(* IEC 61131-3 sources: avi-aoi-management/server/services/programming/iec61131/golden-st/valid, 35 files *)

(* ---- v01-probe-fb.st ---- *)
FUNCTION_BLOCK FB_Light
VAR_INPUT
  Enable : BOOL;
END_VAR
VAR_OUTPUT
  Red : BOOL;
END_VAR
VAR
  T1 : TON;
END_VAR
Red := Enable;
END_FUNCTION_BLOCK

(* ---- v11-fb-in-out-temp-instance.st ---- *)
FUNCTION_BLOCK FB_Accumulate
VAR_INPUT
    Add    : REAL;
    Enable : BOOL;
END_VAR
VAR_IN_OUT
    Total : REAL;
END_VAR
VAR_OUTPUT
    Overflow : BOOL;
END_VAR
VAR_TEMP
    Tmp : REAL;
END_VAR
VAR CONSTANT
    LIMIT_MAX : REAL := 1.0E6;
END_VAR
    IF Enable THEN
        Tmp := Total + Add;
        Overflow := Tmp > LIMIT_MAX;
        IF NOT Overflow THEN
            Total := Tmp;
        END_IF;
    END_IF;
END_FUNCTION_BLOCK

PROGRAM Main
VAR
    Acc     : FB_Accumulate;
    Energy  : REAL;
    Alarm   : BOOL;
END_VAR
    Acc(Add := 0.5, Enable := TRUE, Total := Energy);
    Alarm := Acc.Overflow;
END_PROGRAM

(* ---- v23-traffic-light-fb-timer-array.st ---- *)
FUNCTION_BLOCK FB_TrafficLight
VAR_INPUT
    Enable : BOOL;
END_VAR
VAR_OUTPUT
    Red    : BOOL;
    Yellow : BOOL;
    Green  : BOOL;
END_VAR
VAR
    Phase  : INT := 0;
    Timers : ARRAY[0..2] OF TON;
    Times  : ARRAY[0..2] OF TIME := [T#10s, T#3s, T#8s];
END_VAR

IF NOT Enable THEN
    Phase := 0;
    Red := TRUE; Yellow := FALSE; Green := FALSE;
    RETURN;
END_IF;

Timers[Phase](IN := TRUE, PT := Times[Phase]);
IF Timers[Phase].Q THEN
    Timers[Phase](IN := FALSE);
    Phase := (Phase + 1) MOD 3;
END_IF;

Red := Phase = 0;
Green := Phase = 1;
Yellow := Phase = 2;

END_FUNCTION_BLOCK

PROGRAM Crossing
VAR
    Light : FB_TrafficLight;
    Run   : BOOL := TRUE;
    Stop  : BOOL;
END_VAR
Light(Enable := Run);
Stop := Light.Red;
END_PROGRAM

(* ---- v25-std-functions-conversions.st ---- *)
FUNCTION_BLOCK FB_Clamp
VAR_INPUT
    In   : REAL;
    Lo   : REAL := 0.0;
    Hi   : REAL := 100.0;
END_VAR
VAR_OUTPUT
    Out     : REAL;
    Clipped : BOOL;
    Rounded : INT;
END_VAR
    Out := LIMIT(Lo, In, Hi);
    Clipped := Out <> In;
    Rounded := REAL_TO_INT(Out);
    Rounded := TRUNC(Out);
    Out := MAX(Out, INT_TO_REAL(Rounded));
END_FUNCTION_BLOCK

PROGRAM UseClamp
VAR
    Clamp : FB_Clamp;
    Raw   : REAL;
    Value : REAL;
    Warn  : BOOL;
END_VAR
    Clamp(In := Raw, Hi := 80.0, Out => Value, Clipped => Warn);
END_PROGRAM

(* ---- v32-r-edge-f-edge-inputs.st ---- *)
FUNCTION_BLOCK FB_EdgeCounter
VAR_INPUT
    Pulse   : BOOL R_EDGE;
    Release : BOOL F_EDGE;
    Reset   : BOOL;
END_VAR
VAR_OUTPUT
    Rising  : INT;
    Falling : INT;
END_VAR
IF Reset THEN
    Rising := 0;
    Falling := 0;
END_IF;
IF Pulse THEN
    Rising := Rising + 1;
END_IF;
IF Release THEN
    Falling := Falling + 1;
END_IF;
END_FUNCTION_BLOCK

PROGRAM UseEdges
VAR
    Counter : FB_EdgeCounter;
    Sensor  : BOOL;
    Total   : INT;
END_VAR
Counter(Pulse := Sensor, Release := Sensor, Reset := FALSE);
Total := Counter.Rising;
END_PROGRAM

(* ---- v02-probe-cmt.st ---- *)
PROGRAM P
VAR
  a : BOOL;
END_VAR
(* turn on if sensor is on *)
a := TRUE;
END_PROGRAM

(* ---- v03-conveyor-start-stop-ton.st ---- *)
(* Conveyor: Start push-button latches the motor, NC Stop drops it,
   a TON delays the running lamp by 2 s. *)
PROGRAM ConveyorStartStop
VAR_INPUT
    StartPB   : BOOL;          (* NO push-button *)
    StopPB_NC : BOOL := TRUE;  (* NC push-button: FALSE when pressed *)
END_VAR
VAR_OUTPUT
    Motor      : BOOL;
    RunningLmp : BOOL;
END_VAR
VAR
    RunDelay : TON;
END_VAR

Motor := (StartPB OR Motor) AND StopPB_NC;
RunDelay(IN := Motor, PT := T#2s);
RunningLmp := RunDelay.Q;

END_PROGRAM

(* ---- v04-debounce-ton.st ---- *)
PROGRAM DebounceInputSignal
VAR
    RawSignal    : BOOL;             (* noisy field input *)
    DebounceTmr  : TON;              (* standard on-delay timer instance *)
    StableSignal : BOOL;             (* debounced, steady result (output) *)
    DebounceTime : TIME := T#20ms;   (* dwell needed to accept a change *)
END_VAR

(* TON keeps Q low until IN has stayed high past PT (DebounceTime);
   this rejects contact chatter on a mechanical input. *)
DebounceTmr(IN := RawSignal, PT := DebounceTime);
StableSignal := DebounceTmr.Q;

END_PROGRAM

(* ---- v05-moving-average-array-for.st ---- *)
PROGRAM MovingAverage
VAR
    Samples    : ARRAY[0..7] OF REAL;
    WriteIndex : INT := 0;
    Idx        : INT;
    Sum        : REAL := 0.0;
    NewSample  : REAL;
    Average    : REAL;
END_VAR

Samples[WriteIndex] := NewSample;
WriteIndex := WriteIndex + 1;
IF WriteIndex >= 8 THEN
    WriteIndex := 0;
END_IF;

Sum := 0.0;
FOR Idx := 0 TO 7 DO
    Sum := Sum + Samples[Idx];
END_FOR;
Average := Sum / 8.0;

END_PROGRAM

(* ---- v06-case-enum-state-machine.st ---- *)
TYPE
    E_FillState : (Idle, Filling, Settling, Done);
END_TYPE

PROGRAM FillStation
VAR
    State      : E_FillState := Idle;
    StartReq   : BOOL;
    LevelHigh  : BOOL;
    Valve      : BOOL;
    SettleTmr  : TON;
END_VAR

CASE State OF
    Idle:
        Valve := FALSE;
        IF StartReq THEN
            State := Filling;
        END_IF;
    Filling:
        Valve := TRUE;
        IF LevelHigh THEN
            State := E_FillState#Settling;
        END_IF;
    Settling:
        Valve := FALSE;
        SettleTmr(IN := TRUE, PT := T#3s);
        IF SettleTmr.Q THEN
            SettleTmr(IN := FALSE);
            State := Done;
        END_IF;
    Done:
        IF NOT StartReq THEN
            State := Idle;
        END_IF;
END_CASE;

END_PROGRAM

(* ---- v07-case-int-ranges-else.st ---- *)
PROGRAM SpeedSelector
VAR
    Mode     : INT;
    SpeedSet : REAL;
    Fault    : BOOL;
END_VAR

CASE Mode OF
    0:
        SpeedSet := 0.0;
    1, 2:
        SpeedSet := 25.0;
    3..5:
        SpeedSet := 50.0 + INT_TO_REAL(Mode) * 5.0;
ELSE
    SpeedSet := 0.0;
    Fault := TRUE;
END_CASE

END_PROGRAM

(* ---- v08-while-exit.st ---- *)
PROGRAM FindFirstEmpty
VAR
    Slots     : ARRAY[1..10] OF BOOL;
    I         : INT;
    FirstFree : INT := -1;
END_VAR

I := 1;
WHILE I <= 10 DO
    IF NOT Slots[I] THEN
        FirstFree := I;
        EXIT;
    END_IF;
    I := I + 1;
END_WHILE;

END_PROGRAM

(* ---- v09-repeat-until.st ---- *)
PROGRAM ShiftRegister
VAR
    Reg   : ARRAY[0..4] OF INT;
    K     : INT;
    Input : INT;
END_VAR

K := 4;
REPEAT
    Reg[K] := Reg[K - 1];
    K := K - 1;
UNTIL K = 0
END_REPEAT;
Reg[0] := Input;

END_PROGRAM

(* ---- v10-function-var-input.st ---- *)
FUNCTION Scale : REAL
VAR_INPUT
    Raw    : INT;
    RawMax : INT;
    EngMax : REAL;
END_VAR
    IF RawMax <= 0 THEN
        Scale := 0.0;
        RETURN;
    END_IF;
    Scale := INT_TO_REAL(Raw) / INT_TO_REAL(RawMax) * EngMax;
END_FUNCTION

PROGRAM Main
VAR
    AnalogIn : INT;
    Pressure : REAL;
END_VAR
    Pressure := Scale(Raw := AnalogIn, RawMax := 27648, EngMax := 10.0);
    Pressure := Scale(AnalogIn, 27648, 16.0);
END_PROGRAM

(* ---- v12-ctu-rtrig-batch.st ---- *)
PROGRAM BatchCounter
VAR
    PartSensor : BOOL;
    ResetPB    : BOOL;
    Edge       : R_TRIG;
    Counter    : CTU;
    BatchDone  : BOOL;
    Count      : INT;
END_VAR

Edge(CLK := PartSensor);
Counter(CU := Edge.Q, R := ResetPB, PV := 50);
BatchDone := Counter.Q;
Count := Counter.CV;

END_PROGRAM

(* ---- v13-ctud-ctd.st ---- *)
PROGRAM BufferLevel
VAR
    InSensor  : BOOL;
    OutSensor : BOOL;
    Clear     : BOOL;
    Load      : BOOL;
    Level     : CTUD;
    Remaining : CTD;
    Full      : BOOL;
    Empty     : BOOL;
    Parts     : INT;
END_VAR

Level(CU := InSensor, CD := OutSensor, R := Clear, LD := FALSE, PV := 20);
Full := Level.QU;
Empty := Level.QD;
Parts := Level.CV;
Remaining(CD := OutSensor, LD := Load, PV := 100);
IF Remaining.Q THEN
    Load := TRUE;
END_IF;

END_PROGRAM

(* ---- v14-sr-rs-ftrig.st ---- *)
PROGRAM Latches
VAR
    SetBtn    : BOOL;
    ResetBtn  : BOOL;
    Released  : F_TRIG;
    PumpLatch : SR;
    FanLatch  : RS;
    Pump      : BOOL;
    Fan       : BOOL;
END_VAR

Released(CLK := SetBtn);
PumpLatch(S1 := SetBtn, R := ResetBtn);
FanLatch(S := Released.Q, R1 := ResetBtn);
Pump := PumpLatch.Q1;
Fan := FanLatch.Q1;

END_PROGRAM

(* ---- v15-struct-members.st ---- *)
TYPE
    ST_Axis : STRUCT
        Position : REAL;
        Velocity : REAL;
        Homed    : BOOL;
    END_STRUCT;
    ST_Cell : STRUCT
        AxisX : ST_Axis;
        AxisY : ST_Axis;
        Name  : STRING[32];
    END_STRUCT;
END_TYPE

PROGRAM CellStatus
VAR
    Cell     : ST_Cell;
    AllHomed : BOOL;
    Dist     : REAL;
END_VAR

AllHomed := Cell.AxisX.Homed AND Cell.AxisY.Homed;
Dist := SQRT(Cell.AxisX.Position * Cell.AxisX.Position + Cell.AxisY.Position ** 2.0);
Cell.Name := 'Cell A';

END_PROGRAM

(* ---- v16-comments-with-keywords.st ---- *)
// if this line were code it would be broken: IF x THEN
(* Multi-line comment mentioning for, while, repeat and END_IF / END_FOR
   and even an unbalanced VAR or two: VAR VAR VAR *)
PROGRAM CommentTorture
VAR
    Lamp  : BOOL;   // turn on if the door is open
    Door  : BOOL;   (* while door open, for safety keep lamp on *)
    Label : STRING := 'IF Door THEN END_WHILE (* not a comment *)';
END_VAR
/* block comment: FOR i := 1 TO 10 DO */
IF Door THEN   // for the operator
    Lamp := TRUE;  (* end_if would go here if *)
ELSE
    Lamp := FALSE;
END_IF;
Label := 'it$'s $'quoted$' and // not a comment';
END_PROGRAM

(* ---- v17-global-external-retain.st ---- *)
VAR_GLOBAL
    gMachineReady : BOOL;
    gCycleCount   : DINT;
END_VAR

PROGRAM Cycle
VAR_EXTERNAL
    gMachineReady : BOOL;
    gCycleCount   : DINT;
END_VAR
VAR RETAIN
    TotalCycles : DINT;
END_VAR
VAR CONSTANT
    MAX_CYCLES : DINT := 1000000;
END_VAR
VAR
    CycleStart : BOOL;
    Edge       : R_TRIG;
END_VAR

Edge(CLK := CycleStart AND gMachineReady);
IF Edge.Q AND (TotalCycles < MAX_CYCLES) THEN
    TotalCycles := TotalCycles + 1;
    gCycleCount := TotalCycles;
END_IF;

END_PROGRAM

(* ---- v18-typed-literals.st ---- *)
PROGRAM Literals
VAR
    Mask     : WORD := 16#00FF;
    Bits     : BYTE := 2#1010_0101;
    Oct      : INT := 8#17;
    Small    : INT := INT#5;
    Big      : DINT := 1_000_000;
    Sci      : LREAL := 1.5E-3;
    Neg      : INT := -42;
    Dwell    : TIME := T#1h2m3s;
    Short    : TIME := TIME#500ms;
    Frac     : TIME := T#1.5s;
    Day      : DATE := D#2024-01-31;
    Clock    : TOD := TOD#12:30:00;
    Stamp    : DT := DT#2024-01-31-08:15:00;
    Flag     : BOOL := BOOL#TRUE;
    Masked   : WORD;
END_VAR

Masked := Mask AND 16#0F0F;
IF Dwell > T#1h THEN
    Flag := FALSE;
END_IF;

END_PROGRAM

(* ---- v19-direct-addresses.st ---- *)
PROGRAM IoMapping
VAR
    StartBtn AT %IX0.0 : BOOL;
    StopBtn  AT %IX0.1 : BOOL;
    Motor    AT %QX0.0 : BOOL;
    Speed    AT %IW0   : INT;
    SpeedOut AT %QW0   : INT;
END_VAR

Motor := StartBtn AND NOT StopBtn;
SpeedOut := Speed;
%QX0.1 := Motor;
%MW10 := Speed / 2;

END_PROGRAM

(* ---- v20-expressions-operators.st ---- *)
PROGRAM Expressions
VAR
    A, B, C : BOOL;
    X, Y    : INT;
    R       : REAL;
    Res     : BOOL;
    Parity  : INT;
END_VAR

Res := (A AND B) OR (NOT C XOR A) & (X <> Y);
Res := (X >= 10) AND (Y <= -3) OR (X = Y) AND NOT (X > Y OR X < Y);
Parity := X MOD 2;
R := INT_TO_REAL(X) ** 2.0 + INT_TO_REAL(Y) / 3.0 - 1.0;
X := -(Y * 4) + ABS(Y) - MAX(X, Y) + MIN(X, 0) + LIMIT(0, Y, 100);
Res := SEL(A, B, C);

END_PROGRAM

(* ---- v21-fb-output-binding.st ---- *)
PROGRAM OutputBinding
VAR
    Go       : BOOL;
    Tmr      : TON;
    Done     : BOOL;
    Elapsed  : TIME;
    Pulse    : TP;
    OffDelay : TOF;
    PulseOut : BOOL;
    Hold     : BOOL;
END_VAR

Tmr(IN := Go, PT := T#2s, Q => Done, ET => Elapsed);
Pulse(IN := Done, PT := T#500ms, Q => PulseOut);
OffDelay(IN := Go, PT := T#5s);
Hold := OffDelay.Q AND NOT Pulse.Q;

END_PROGRAM

(* ---- v22-nested-if-for-by.st ---- *)
PROGRAM Nested
VAR
    Data  : ARRAY[1..20] OF INT;
    I     : INT;
    Pos   : INT;
    Neg   : INT;
    Zero  : INT;
END_VAR

Pos := 0; Neg := 0; Zero := 0;
FOR I := 20 TO 1 BY -1 DO
    IF Data[I] > 0 THEN
        Pos := Pos + 1;
    ELSIF Data[I] < 0 THEN
        Neg := Neg + 1;
        IF Neg > 5 THEN
            EXIT;
        END_IF;
    ELSE
        Zero := Zero + 1;
    END_IF;
END_FOR;

END_PROGRAM

(* ---- v24-strings-bits-multidim.st ---- *)
PROGRAM StringsAndBits
VAR
    Status  : WORD;
    Ready   : BOOL;
    Msg     : STRING(80);
    Prefix  : STRING := 'Line';
    Grid    : ARRAY[1..3, 1..4] OF INT;
    MsgLen  : INT;
    R, C    : INT;
END_VAR

Ready := Status.3;
Status.0 := TRUE;
Msg := CONCAT(Prefix, ' 1 ready');
MsgLen := LEN(Msg);
FOR R := 1 TO 3 DO
    FOR C := 1 TO 4 DO
        Grid[R, C] := R * 10 + C;
    END_FOR;
END_FOR;

END_PROGRAM

(* ---- v26-unbounded-while-lint-only.st ---- *)
(* Syntactically valid; the SAFETY linter (not the parser) flags the unbounded loop. *)
PROGRAM ConveyorPoll
VAR
    SensorInput : BOOL;
    MotorRun    : BOOL;
END_VAR

WHILE TRUE DO
    MotorRun := SensorInput;
END_WHILE;

END_PROGRAM

(* ---- v27-time-date-functions.st ---- *)
PROGRAM TimeArithmetic
VAR
    Dwell     : TIME := T#2s;
    Extra     : TIME := T#500ms;
    Total     : TIME;
    Diff      : TIME;
    Scaled    : TIME;
    Half      : TIME;
    ShiftTod  : TOD := TOD#06:00:00;
    NowTod    : TOD := TOD#14:30:00;
    LaterTod  : TOD;
    EarlyTod  : TOD;
    Stamp     : DT := DT#2024-01-31-08:15:00;
    Stamp2    : DT;
    Stamp3    : DT;
    Day1      : DATE := D#2024-01-01;
    Day2      : DATE := D#2024-02-01;
    DaySpan   : TIME;
    TodSpan   : TIME;
    DtSpan    : TIME;
    Joined    : DT;
END_VAR

Total := ADD_TIME(Dwell, Extra);
Diff := SUB_TIME(Dwell, Extra);
Scaled := MULTIME(Dwell, 3);
Half := DIVTIME(Dwell, 2);
LaterTod := ADD_TOD_TIME(ShiftTod, T#8h);
EarlyTod := SUB_TOD_TIME(NowTod, T#30m);
TodSpan := SUB_TOD_TOD(NowTod, ShiftTod);
Stamp2 := ADD_DT_TIME(Stamp, T#1h);
Stamp3 := SUB_DT_TIME(Stamp, T#15m);
DtSpan := SUB_DT_DT(Stamp2, Stamp);
DaySpan := SUB_DATE_DATE(Day2, Day1);
Joined := CONCAT_DATE_TOD(Day1, ShiftTod);

END_PROGRAM

(* ---- v28-long-conversions-bcd.st ---- *)
PROGRAM Conversions
VAR
    Stamp    : DATE_AND_TIME := DT#2024-01-31-08:15:00;
    ClockTod : TIME_OF_DAY;
    OnlyDay  : DATE;
    Raw      : WORD := 16#0123;
    Value    : INT;
    Back     : WORD;
    R        : REAL := 12.7;
    I        : DINT;
    Text     : STRING;
    B        : BOOL;
END_VAR

ClockTod := DATE_AND_TIME_TO_TIME_OF_DAY(Stamp);
OnlyDay := DATE_AND_TIME_TO_DATE(Stamp);
ClockTod := DT_TO_TOD(Stamp);
Value := WORD_BCD_TO_INT(Raw);
Value := BCD_TO_INT(Raw);
Back := INT_TO_BCD(Value);
I := REAL_TO_DINT(R);
I := TRUNC(R);
Text := INT_TO_STRING(Value);
B := INT_TO_BOOL(Value);

END_PROGRAM

(* ---- v29-numeric-selection-shift.st ---- *)
PROGRAM NumericSelectShift
VAR
    X, Y, Z  : REAL;
    A, B     : INT;
    W        : WORD := 16#00F0;
    G        : BOOL;
    K        : INT := 1;
    Cmp      : BOOL;
END_VAR

X := ABS(Y) + SQRT(Z) + LN(Z) + LOG(Z) + EXP(Y);
X := SIN(Y) + COS(Y) + TAN(Y) + ASIN(Z) + ACOS(Z) + ATAN(Z);
X := EXPT(Y, 2.0);
A := ADD(A, B, 3);
A := SUB(A, B);
A := MUL(A, B);
A := DIV(A, 2);
A := MOVE(B);
A := SEL(G, A, B);
A := MAX(A, B, 7);
A := MIN(A, B);
A := LIMIT(0, A, 100);
A := MUX(K, 10, 20, 30);
W := SHL(W, 2);
W := SHR(W, 1);
W := ROL(W, 4);
W := ROR(W, 4);
Cmp := GT(A, B) OR GE(A, B) OR EQ(A, B) OR LE(A, B) OR LT(A, B) OR NE(A, B);

END_PROGRAM

(* ---- v30-string-functions.st ---- *)
PROGRAM StringFunctions
VAR
    S1   : STRING := 'Line-1 ready';
    S2   : STRING;
    N    : INT;
    P    : INT;
END_VAR

N := LEN(S1);
S2 := LEFT(S1, 4);
S2 := RIGHT(S1, 5);
S2 := MID(S1, 2, 6);
S2 := CONCAT(S2, ' / ', S1);
S2 := INSERT(S1, 'X', 3);
S2 := DELETE(S1, 2, 1);
S2 := REPLACE(S1, 'OK', 2, 7);
P := FIND(S1, 'ready');

END_PROGRAM

(* ---- v31-operator-call-forms.st ---- *)
PROGRAM OperatorCallForms
VAR
    A, B, C : BOOL;
    W1, W2  : WORD;
    N       : INT := 17;
    R       : INT;
END_VAR

R := MOD(N, 5);
C := AND(A, B);
C := OR(A, B, C);
C := XOR(A, B);
C := NOT(A);
W1 := AND(W1, W2);
C := A AND (B OR NOT C);

END_PROGRAM

(* ---- v33-comment-mentions-open-marker.st ---- *)
(* To start a comment write (* and close it with the matching marker *)
PROGRAM CommentMarkerText
VAR
    Lamp : BOOL;  (* note: "(*" alone is just text here *)
END_VAR
Lamp := TRUE;
END_PROGRAM

(* ---- v34-comment-mentions-marker-then-string-close.st ---- *)
(* Reviewer repro (fix round 2): this comment mentions (* in its text and is closed here *)
PROGRAM CommentThenStringMarker
VAR
    Hint  : STRING := 'end a comment with *)';
    Lamp  : BOOL;
    Count : INT;
END_VAR

Lamp := TRUE;
Count := Count + 1;
Hint := 'end a comment with *)';

END_PROGRAM

(* ---- v35-standard-conversion-names.st ---- *)
PROGRAM StandardConversions
VAR
    Stamp   : DATE_AND_TIME := DT#2024-01-31-08:15:00;
    Clock   : TIME_OF_DAY;
    Count   : DINT := 42;
    Ratio   : REAL;
    Raw     : WORD := 16#0042;
    Small   : INT;
    Packed  : WORD;
    Big     : LREAL := 3.9;
    Whole   : DINT;
END_VAR

Clock := DATE_AND_TIME_TO_TIME_OF_DAY(Stamp);
Ratio := DINT_TO_REAL(Count) / 10.0;
Small := WORD_BCD_TO_INT(Raw);
Packed := INT_TO_BCD_WORD(Small);
Whole := LREAL_TRUNC_DINT(Big);
Small := TO_INT(Ratio);
Ratio := LREAL_TO_REAL(Big);

END_PROGRAM
